(* IEC 61131-3 sources: Test-Git_ESME26/TestProgettoESME_26.fbsproj/PacDriveLib Migration/Motion/MultiCam/PDL_FB_MultiCam.fb.st^/Check, 4 files *)

(* ---- CheckCamData.meth.st ---- *)
METHOD CheckCamData : BOOL
VAR_INPUT
END_VAR

//return TRUE: data is valid
CheckCamData := TRUE;

//check cam data
IF iq_stMultiCamData.diNumberOfCamPoints <= 0 OR iq_stMultiCamData.diNumberOfCamPoints > UPPER_BOUND(iq_stMultiCamData.astCamPoint, 1) THEN

	SetDiagOutput(	i_etDiag	:= GD.ET_Diag.InputParameterInvalid,
					i_etDiagExt := PDL_ET_DiagExt.NumberOfCamPointsRange,
					i_sMsg		:= SE_CTBX.FC_MultiConcat(	i_sString1 := '0 < ST_MultiCam.diNumberOfCamPoints <= ',
															i_sString2 := DINT_TO_STRING( UPPER_BOUND(iq_stMultiCamData.astCamPoint, 1) ),
															i_sString3 := ' , Current: ',
															i_sString4 := DINT_TO_STRING(iq_stMultiCamData.diNumberOfCamPoints) )
					);

	q_xSynActive		:= FALSE;
	q_xXLowEnd			:= FALSE;
	q_xXHighEnd			:= FALSE;
	iq_xNewCam			:= FALSE;
	iq_xInstantNewCam	:= FALSE;

	etState := ET_MulticamState.controllerStop;

	CheckCamData := FALSE;

END_IF

(* ---- InputParameterCheck.meth.st ---- *)
METHOD PRIVATE InputParameterCheck : BOOL
VAR_INPUT
	i_xCheckWsParam			: BOOL;
	i_xCheckStartPosParam	: BOOL;
	i_xCheckStopPosParam	: BOOL;
END_VAR

VAR
	lrMaxAcc	: LREAL := 0;
	lrMaxVel	: LREAL := 0;
END_VAR

InputParameterCheck := FALSE;

//if IF_DriveConfig is not available -> limits are NOT checked
IF ifDriveConfig <> 0 THEN
	lrMaxAcc := ifDriveConfig.MaxAcc;
	lrMaxVel := ifDriveConfig.MaxVel;
END_IF

IF  ABS(i_lrWsVel) > lrMaxVel AND lrMaxVel <> 0  AND i_xCheckWsParam THEN
		SetDiagOutput(	i_etDiag	:= GD.ET_Diag.InputParameterInvalid,
						i_etDiagExt := PDL_ET_DiagExt.VelRange,
						i_sMsg		:= SE_CTBX.FC_MultiConcat(	i_sString1 := 'i_lrWsVel',
																i_sString2 := ' <= ',
																i_sString3 := TO_STRING(lrMaxVel),
																i_sString4 := '') );

ELSIF (i_lrWsAcc <= 0 OR (i_lrWsAcc > lrMaxAcc AND lrMaxAcc <> 0)) AND i_xCheckWsParam THEN
		SetDiagOutput(	i_etDiag	:= GD.ET_Diag.InputParameterInvalid,
						i_etDiagExt := PDL_ET_DiagExt.AccRange,
						i_sMsg		:= SE_CTBX.FC_MultiConcat(	i_sString1 := '0.0 < ',
																i_sString2 := 'i_lrWsAcc',
																i_sString3 := ' <= ',
																i_sString4 := TO_STRING(lrMaxAcc) ));

ELSIF (i_lrWsJerk <= 0.0 ) AND i_xCheckWsParam THEN
		SetDiagOutput(	i_etDiag	:= GD.ET_Diag.InputParameterInvalid,
						i_etDiagExt := PDL_ET_DiagExt.JerkRange,
						i_sMsg		:= '0.0 < i_lrWsJerk ');

ELSIF iq_stExt.xStartPositionSelect AND  (ABS(iq_stExt.lrStartVelocity) > lrMaxVel AND lrMaxVel <> 0) AND i_xCheckStartPosParam THEN
 		SetDiagOutput(	i_etDiag	:= GD.ET_Diag.InputParameterInvalid,
 						i_etDiagExt := PDL_ET_DiagExt.VelRange,
 						i_sMsg		:= SE_CTBX.FC_MultiConcat(	i_sString1 := 'iq_stExt.lrStartVelocity',
																i_sString2 := ' <= ',
																i_sString3 := TO_STRING(lrMaxVel),
																i_sString4 := ''));

ELSIF iq_stExt.xStartPositionSelect AND (iq_stExt.lrStartAcceleration <= 0 OR (iq_stExt.lrStartAcceleration > lrMaxAcc AND lrMaxAcc <> 0) ) AND i_xCheckStartPosParam THEN
		SetDiagOutput(	i_etDiag	:= GD.ET_Diag.InputParameterInvalid,
						i_etDiagExt := PDL_ET_DiagExt.AccRange,
						i_sMsg		:= SE_CTBX.FC_MultiConcat(	i_sString1 := '0.0 < ',
																i_sString2 := 'iq_stExt.lrStartAcceleration',
																i_sString3 := ' <= ',
																i_sString4 := TO_STRING(lrMaxAcc) ));

ELSIF iq_stExt.xStartPositionSelect AND (iq_stExt.lrStartDeceleration <= 0 OR (iq_stExt.lrStartDeceleration > lrMaxAcc AND lrMaxAcc <> 0) ) AND i_xCheckStartPosParam THEN
		SetDiagOutput(	i_etDiag	:= GD.ET_Diag.InputParameterInvalid,
						i_etDiagExt := PDL_ET_DiagExt.DecRange,
						i_sMsg		:= SE_CTBX.FC_MultiConcat(	i_sString1 := '0.0 < ',
																i_sString2 := 'iq_stExt.lrStartDeceleration',
																i_sString3 := ' <= ',
																i_sString4 := TO_STRING(lrMaxAcc) ));

ELSIF iq_stExt.xStartPositionSelect AND (iq_stExt.lrStartJerk <= 0.0 ) AND i_xCheckStartPosParam THEN
		SetDiagOutput(	i_etDiag	:= GD.ET_Diag.InputParameterInvalid,
						i_etDiagExt := PDL_ET_DiagExt.JerkRange,
						i_sMsg		:= '0.0 < iq_stExt.lrStartJerk');

ELSIF iq_stExt.xStopPositionSelect AND (ABS(iq_stExt.lrStopVelocity) > lrMaxVel AND lrMaxVel <> 0) AND i_xCheckStopPosParam THEN
 		SetDiagOutput(	i_etDiag	:= GD.ET_Diag.InputParameterInvalid,
 						i_etDiagExt := PDL_ET_DiagExt.VelRange,
 						i_sMsg		:= SE_CTBX.FC_MultiConcat(	i_sString1 := 'iq_stExt.lrStopVelocity',
																i_sString2 := ' <= ',
																i_sString3 := TO_STRING(lrMaxVel),
																i_sString4 := ''));

ELSIF iq_stExt.xStopPositionSelect AND (iq_stExt.lrStopAcceleration <= 0 OR (iq_stExt.lrStopAcceleration > lrMaxAcc AND lrMaxAcc <> 0) ) AND i_xCheckStopPosParam THEN
		SetDiagOutput(	i_etDiag	:= GD.ET_Diag.InputParameterInvalid,
						i_etDiagExt := PDL_ET_DiagExt.AccRange,
						i_sMsg		:= SE_CTBX.FC_MultiConcat(	i_sString1 := '0.0 < ',
																i_sString2 := 'iq_stExt.lrStopAcceleration',
																i_sString3 := ' <= ',
																i_sString4 := TO_STRING(lrMaxAcc) ));

ELSIF iq_stExt.xStopPositionSelect AND (iq_stExt.lrStopDeceleration <= 0 OR (iq_stExt.lrStopDeceleration > lrMaxAcc AND lrMaxAcc <> 0)) AND i_xCheckStopPosParam THEN
		SetDiagOutput(	i_etDiag	:= GD.ET_Diag.InputParameterInvalid,
						i_etDiagExt := PDL_ET_DiagExt.DecRange,
						i_sMsg		:= SE_CTBX.FC_MultiConcat(	i_sString1 := '0.0 < ',
																i_sString2 := 'iq_stExt.lrStopDeceleration',
																i_sString3 := ' <= ',
																i_sString4 := TO_STRING(lrMaxAcc) ));

ELSIF iq_stExt.xStopPositionSelect AND (iq_stExt.lrStopJerk <= 0.0 ) AND i_xCheckStopPosParam THEN
		SetDiagOutput(	i_etDiag	:= GD.ET_Diag.InputParameterInvalid,
						i_etDiagExt := PDL_ET_DiagExt.JerkRange,
						i_sMsg		:= '0.0 < iq_stExt.lrStopJerk');

ELSE
	InputParameterCheck := TRUE;
END_IF

(* ---- MasterMovedCheck.meth.st ---- *)
METHOD PRIVATE MasterMovedCheck : BOOL
VAR_INPUT
END_VAR

MasterMovedCheck := FALSE;

//check master position again...
xSuccess :=  GetCamPositionOfSlave( i_xCheckModulo 		:= FALSE,
									q_lrSlavePosition 	=> lrYStart2 );

IF NOT xSuccess THEN
	RETURN;
END_IF

//...and compare to first position
IF ABS(lrYStart - lrYStart2) > 1.0 THEN
	q_xReady := FALSE;
	SetDiagOutput(	i_etDiag	:= GD.ET_Diag.WarmStartConditionInvalid,
					i_etDiagExt := PDL_ET_DiagExt.MasterMoved,
					i_sMsg		:= '');
	q_xInWSWindow := FALSE;

	etState := ET_MulticamState.controllerStop;
ELSE
	//no master movement detected -> success
	MasterMovedCheck := TRUE;

END_IF

(* ---- YEqualCheck.meth.st ---- *)
METHOD INTERNAL YEqualCheck : BOOL

VAR_INPUT
	i_lrYValueOldCam	: LREAL;
	i_lrYValueNewCam	: LREAL;
	i_lrPeriod			: LREAL;
	i_lrAccuracy		: LREAL;
END_VAR

VAR
	lrDiff				: LREAL;
	lrPeriode			: LREAL;
END_VAR

YEqualCheck := TRUE;

lrDiff:=	ABS(i_lrYValueOldCam - i_lrYValueNewCam);
lrPeriode:= ABS(i_lrPeriod);

IF lrPeriode > CMT.GCL.Gc_lrZeroTolerance THEN
	lrDiff:= MATH.fmod(lrX:= lrDiff, lrM:= lrPeriode);
END_IF

IF 	lrDiff > i_lrAccuracy THEN
	YEqualCheck:= FALSE;
END_IF
